// TIA Portal V17 export
// export: Created 2026-11-20T13:38:29.1107445Z, ExportSetting None, DisplayName Totally Integrated Automation Portal, DisplayVersion V17 Update 9, DisplayName TIA Portal Openness, DisplayVersion V17 Update 9, DisplayName TIA Portal Teamcenter Gateway, DisplayVersion V17 Update 9, DisplayName TIA Portal Version Control Interface, DisplayVersion V17 Update 9, DisplayName Simotion SCOUT TIA, DisplayVersion 5.4.3.0, DisplayName TIA Portal Test Suite Advanced, DisplayVersion V17 Update 1, DisplayName SIMOCODE ES, DisplayVersion V17 Update 8, DisplayName SINAMICS Startdrive Advanced, DisplayVersion V17 SP2, DisplayName SINAMICS DCC, DisplayVersion V17 Update 1, DisplayName SINAMICS Startdrive G110M, G120, G120C, G120D, G120P, G115D, DisplayVersion V17 SP2, DisplayName SINAMICS Startdrive G130, G150, S120, S150, SINAMICS MV, S210, DisplayVersion V17 SP2, DisplayName SIRIUS Safety ES, DisplayVersion V17 Update 8, DisplayName SIRIUS Soft Starter ES, DisplayVersion V17 Update 8, DisplayName STEP 7 Professional, DisplayVersion V17 Update 9, DisplayName SINUMERIK ONE STEP 7 Toolbox, DisplayVersion V17 Update 12, DisplayName SINUMERIK ONE PLC Basic Program Plus, DisplayVersion V17 Update 12, DisplayName SIMATIC Energy Suite, DisplayVersion V17 Update 4, DisplayName STEP 7 CFC, DisplayVersion V17 Update 1, DisplayName SINUMERIK 840D sl STEP 7 Toolbox, DisplayVersion V17 Update 12, DisplayName SINUMERIK MC STEP 7 Toolbox, DisplayVersion V17 Update 12, DisplayName STEP 7 Safety, DisplayVersion V17 Update 6, DisplayName WinCC Professional, DisplayVersion V17 Update 9, DisplayName SIMATIC Visualization Architect, DisplayVersion V17 Update 9, DisplayName SINUMERIK Integrate Create MyHMI /WinCC, DisplayVersion V17
FUNCTION_BLOCK "MCP_RC_FB"   // FB1, SCL
{ S7_Optimized_Access := 'TRUE' }
// stored: MemoryReserve 100, SetENOAutomatically false
   VAR_INPUT
      Start : Bool;
   END_VAR
   VAR_OUTPUT
      Run : Bool;
   END_VAR
   VAR
      Total : Int;
   END_VAR
BEGIN

   #Run := #Start AND "MCP_RC_DB".Status.Ready;
   #Total := "MCP_RC_FC"("A" := #Total, "B" := "MCP_RC_DB".Count);
END_FUNCTION_BLOCK
